TYPE ST_Error :
STRUCT
	b_Active				: BOOL;
	b_memo				: BOOL;
	(*e_Description			: E_ErrorList;*)
	iErNum				: INT;
END_STRUCT
END_TYPE

(* stored: Version 1.1.0.1, ProductVersion 3.1.4024.13
   DUT ST_Error: Id {cdd7197c-8a8a-4300-8532-ed3ea601df7a} *)
